TYPE coffee :
STRUCT
	
price			: REAL;
name			: STRING;
ingredients		: STRING;


END_STRUCT
END_TYPE

(* stored: Version 1.1.0.1
   DUT coffee: Id {94d45191-96d5-4f79-b3b6-aad804f7ddbd} *)
